Fanuc KAREL source: KT00888.KL

PROGRAM KT00888
%NOLOCKGROUP
VAR
  P1: POSITION
  P2: POSITION
  OUT: POSITION
BEGIN
  OUT = INV(P1)
END KT00888
